(* Logix 5000 project; controller R400_500_XLS vendor 1 type 14 code 216 rev 31.11; software revision 31.01; part 25 of 32 *)
(* tags used below, declared in another part *)
   Abort1 : DINT;   // Not Used
   Alarm : SINT;   // Wait 3 seconds
   AlarmAcked : BOOL;   // Alarm has been acked
   bAlrm : BOOL[64];
   CycExcBuffer : UDT_CYCLE;
   DrainNo : DINT;
   DrnSmp : DINT;
   DRYING : DINT;   // Drying id number
   F1rinse : DINT;   // Not Used
   Fill_Sump : DINT;
   Inj_Time : SINT;   // Time based chemical injection steps
   Last_PwWshRnseTtr : DINT;
   M : DINT[5];   // Memory Bits
   ONS_FC11 : DINT;
   ONS_FC13 : DINT;
   PwExcBuffer : UDT_PW;
   RinseExcBuffer : UDT_RINSE;
   Run : DINT;
   SumpWaterVolume : DINT;   // Sump Water Volume 0 =Low 1= High
   Tmr : TIMER[107];
   Trt_PrWsh : DINT;
   Trt_Rinse : DINT;   // Rinse steps
   Trt_Wsh : DINT;
   WASH_1 : DINT;   // Wash 1 id number
   WASH_5 : DINT;   // Wash 5 id number
   WaterSaved : BOOL;   // Water Saved In Sump (Last Final Rinse Water)
   WshExcBuffer : UDT_WASH;
   bPureWaterFillingAuthorization : BOOL;   // Pure Water Filling Authorization Signal
   DrainExtensionTime : DINT;
   I_Shlf_Sw : BOOL;   // Shelf switch
   I_Smp_Lvl_Hgh : BOOL;   // Sump high level switch
   I_Smp_Lvl_Lw : BOOL;   // Sump low level switch
   msg : BOOL[512];
   PreHeatTime : DINT;
   SumpAlarmFillTime : DINT;
   SumpTemp : REAL;   // Sump temperature in °C
   SumpTempToCool : REAL;   // Sump temperature in °C
   tDelayBeforeFillingAuthAlarm : TIMER;
   tPWClosingDelay : TIMER;
   TreatmentPtr : DINT;
   Unit : Hrdwre;   // Unit Configuration
(* MainProgram, continued *)

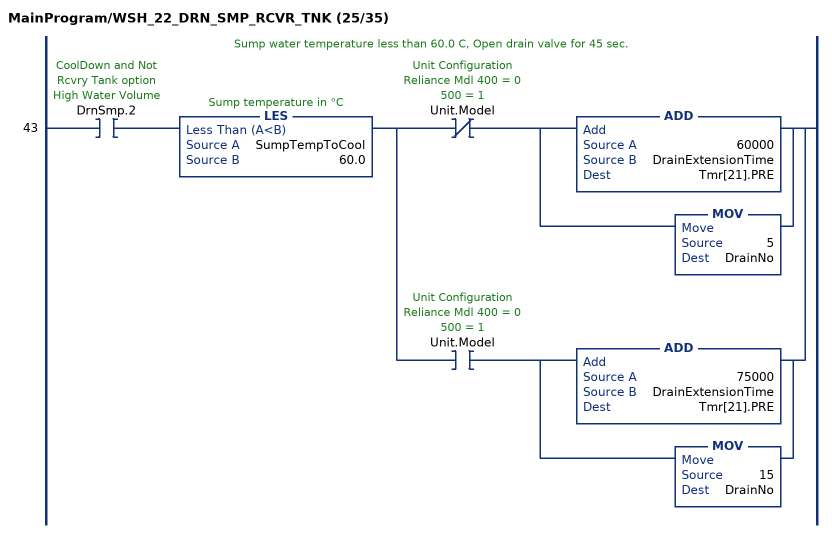
   [picture p501: MainProgram/WSH_22_DRN_SMP_RCVR_TNK rungs 43-43]
   // Sump water temperature less than 60.0 C, Open drain valve for 45 sec.
   43: XIC(DrnSmp.2)LES(SumpTempToCool,60.0)[XIO(Unit.Model) [ADD(60000,DrainExtensionTime,Tmr[21].PRE) ,MOV(5,DrainNo) ] ,XIC(Unit.Model) [ADD(75000,DrainExtensionTime,Tmr[21].PRE) ,MOV(15,DrainNo) ] ];
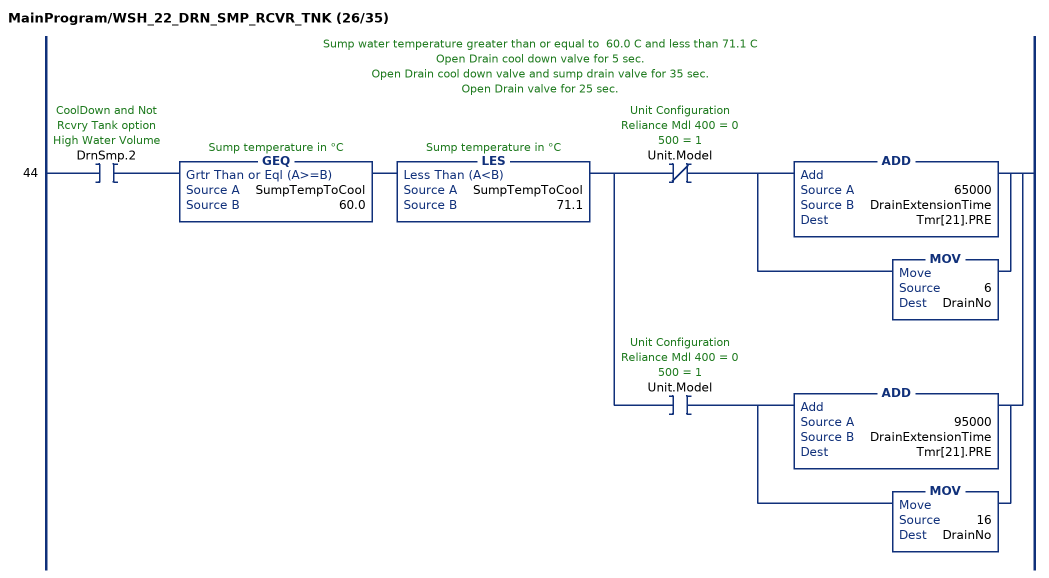
   // Sump water temperature greater than or equal to  60.0 C and less than 71.1 C
   // Open Drain cool down valve for 5 sec.
   // Open Drain cool down valve and sump drain valve for 35 sec.
   // Open Drain valve for 25 sec.
   44: XIC(DrnSmp.2)GEQ(SumpTempToCool,60.0)LES(SumpTempToCool,71.1)[XIO(Unit.Model) [ADD(65000,DrainExtensionTime,Tmr[21].PRE) ,MOV(6,DrainNo) ] ,XIC(Unit.Model) [ADD(95000,DrainExtensionTime,Tmr[21].PRE) ,MOV(16,DrainNo) ] ];
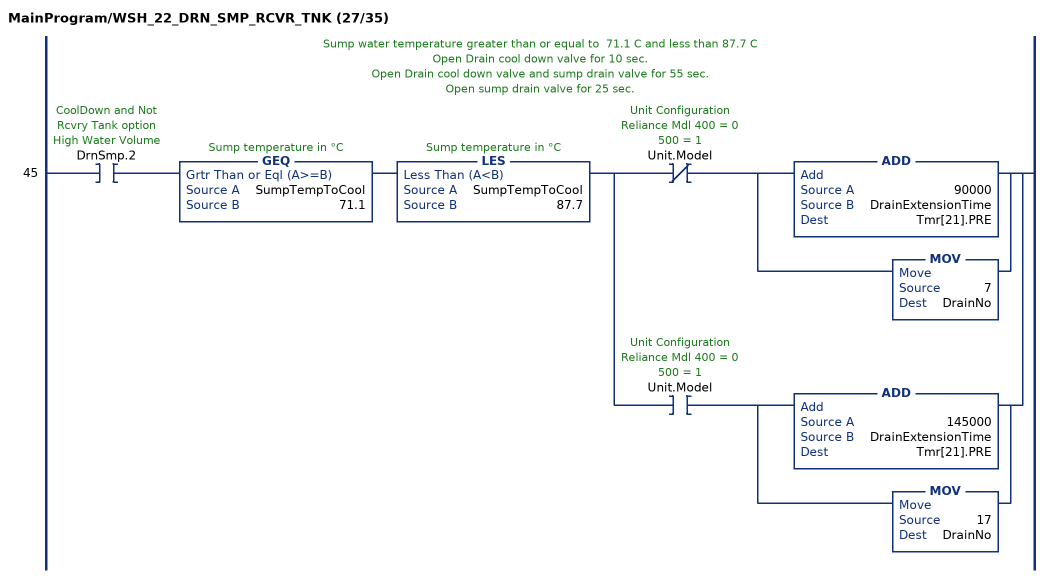
   // Sump water temperature greater than or equal to  71.1 C and less than 87.7 C
   // Open Drain cool down valve for 10 sec.
   // Open Drain cool down valve and sump drain valve for 55 sec.
   // Open sump drain valve for 25 sec.
   45: XIC(DrnSmp.2)GEQ(SumpTempToCool,71.1)LES(SumpTempToCool,87.7)[XIO(Unit.Model) [ADD(90000,DrainExtensionTime,Tmr[21].PRE) ,MOV(7,DrainNo) ] ,XIC(Unit.Model) [ADD(145000,DrainExtensionTime,Tmr[21].PRE) ,MOV(17,DrainNo) ] ];
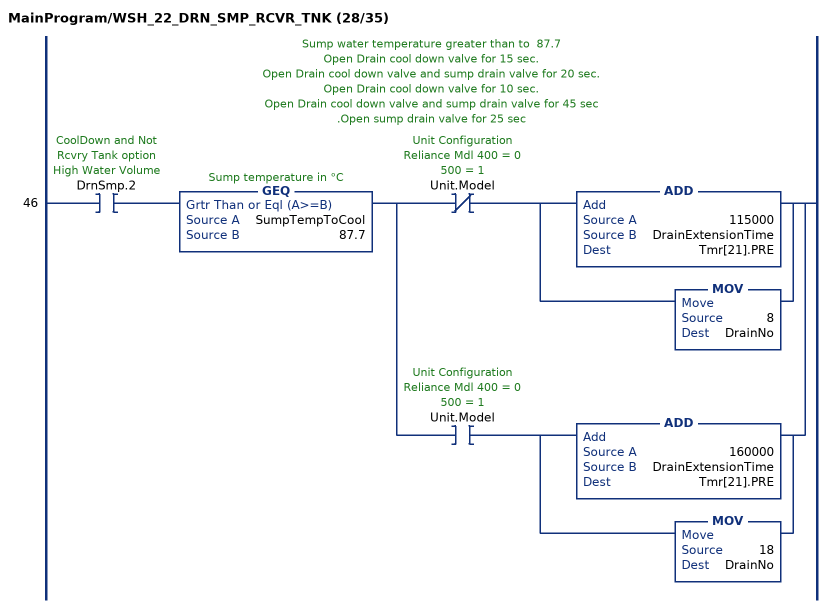
   // Sump water temperature greater than to  87.7
   // Open Drain cool down valve for 15 sec.
   // Open Drain cool down valve and sump drain valve for 20 sec.
   // Open Drain cool down valve for 10 sec.
   // Open Drain cool down valve and sump drain valve for 45 sec
   // .Open sump drain valve for 25 sec
   46: XIC(DrnSmp.2)GEQ(SumpTempToCool,87.7)[XIO(Unit.Model) [ADD(115000,DrainExtensionTime,Tmr[21].PRE) ,MOV(8,DrainNo) ] ,XIC(Unit.Model) [ADD(160000,DrainExtensionTime,Tmr[21].PRE) ,MOV(18,DrainNo) ] ];
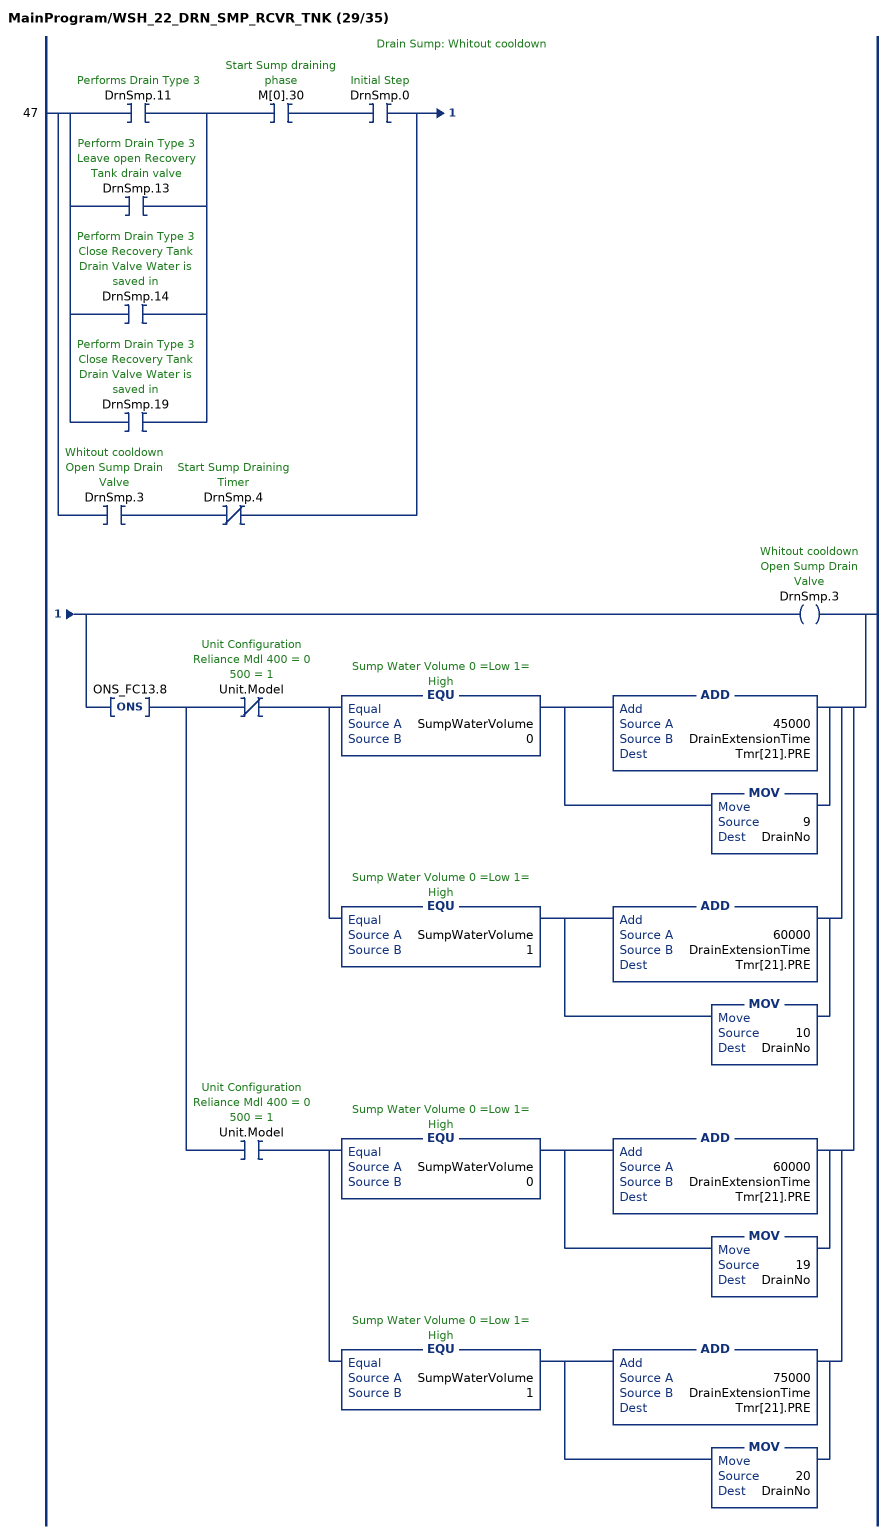
   // Drain Sump: Whitout cooldown
   47: [[XIC(DrnSmp.11) ,XIC(DrnSmp.13) ,XIC(DrnSmp.14) ,XIC(DrnSmp.19) ] XIC(M[0].30) XIC(DrnSmp.0) ,XIC(DrnSmp.3) XIO(DrnSmp.4) ][OTE(DrnSmp.3) ,ONS(ONS_FC13.8) [XIO(Unit.Model) [EQU(SumpWaterVolume,0) [ADD(45000,DrainExtensionTime,Tmr[21].PRE) ,MOV(9,DrainNo) ] ,EQU(SumpWaterVolume,1) [ADD(60000,DrainExtensionTime,Tmr[21].PRE) ,MOV(10,DrainNo) ] ] ,XIC(Unit.Model) [EQU(SumpWaterVolume,0) [ADD(60000,DrainExtensionTime,Tmr[21].PRE) ,MOV(19,DrainNo) ] ,EQU(SumpWaterVolume,1) [ADD(75000,DrainExtensionTime,Tmr[21].PRE) ,MOV(20,DrainNo) ] ] ] ];
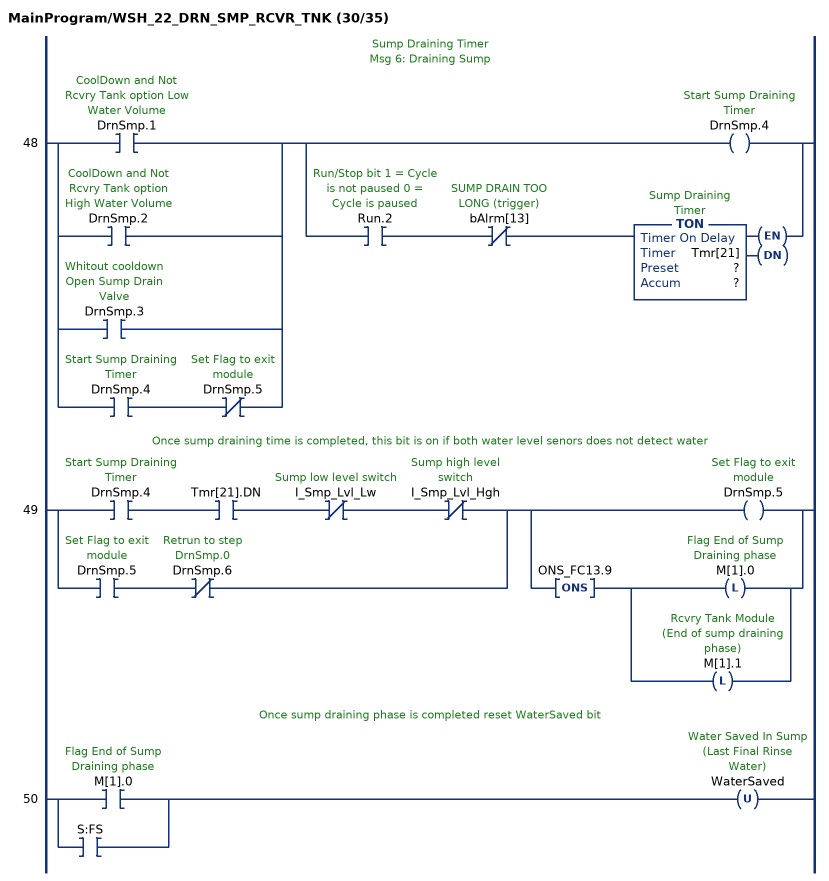
   // Sump Draining Timer
   // Msg 6: Draining Sump
   48: [[XIC(DrnSmp.1) ,XIC(DrnSmp.2) ,XIC(DrnSmp.3) ] ,XIC(DrnSmp.4) XIO(DrnSmp.5) ][OTE(DrnSmp.4) ,XIC(Run.2) XIO(bAlrm[13]) TON(Tmr[21],?,?) ];
   // Once sump draining time is completed, this bit is on if both water level senors does not detect water
   49: [XIC(DrnSmp.4) XIC(Tmr[21].DN) XIO(I_Smp_Lvl_Lw) XIO(I_Smp_Lvl_Hgh) ,XIC(DrnSmp.5) XIO(DrnSmp.6) ][OTE(DrnSmp.5) ,ONS(ONS_FC13.9) [OTL(M[1].0) ,OTL(M[1].1) ] ];
   // Once sump draining phase is completed reset WaterSaved bit
   50: [XIC(M[1].0) ,XIC(S:FS) ]OTU(WaterSaved);
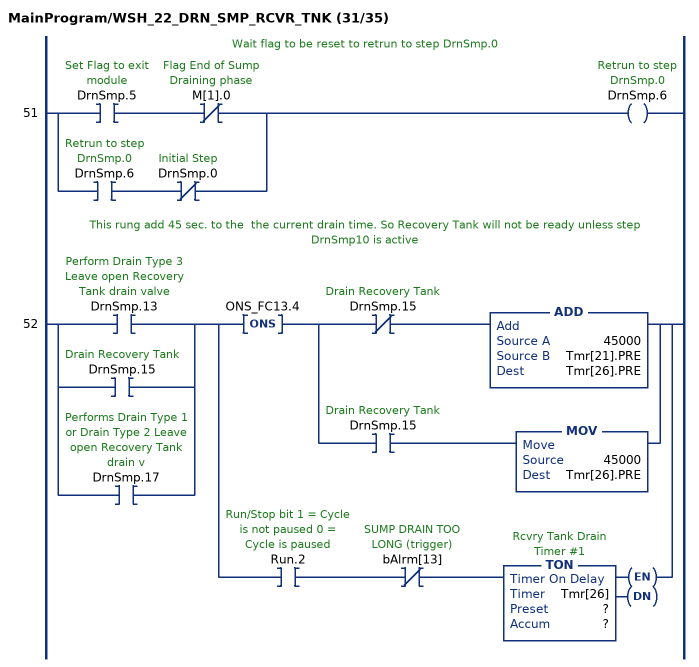
   // Wait flag to be reset to retrun to step DrnSmp.0
   51: [XIC(DrnSmp.5) XIO(M[1].0) ,XIC(DrnSmp.6) XIO(DrnSmp.0) ]OTE(DrnSmp.6);
   // This rung add 45 sec. to the  the current drain time. So Recovery Tank will not be ready unless step DrnSmp10 is active
   52: [XIC(DrnSmp.13) ,XIC(DrnSmp.15) ,XIC(DrnSmp.17) ][ONS(ONS_FC13.4) [XIO(DrnSmp.15) ADD(45000,Tmr[21].PRE,Tmr[26].PRE) ,XIC(DrnSmp.15) MOV(45000,Tmr[26].PRE) ] ,XIC(Run.2) XIO(bAlrm[13]) TON(Tmr[26],?,?) ];
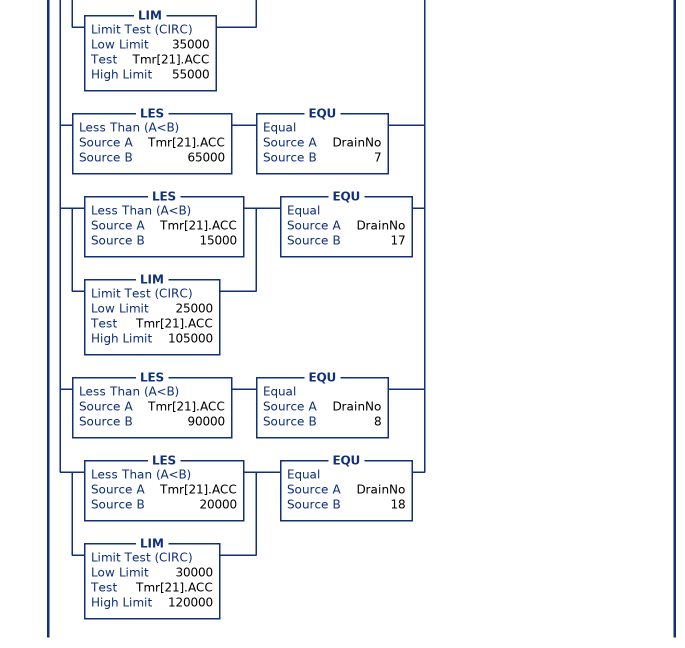
   // Open drain cooldown valve
   53: [LES(Tmr[21].ACC,25000) EQU(DrainNo,2) ,LES(Tmr[21].ACC,35000) EQU(DrainNo,12) ,LES(Tmr[21].ACC,45000) EQU(DrainNo,3) ,[LES(Tmr[21].ACC,15000) ,LIM(25000,Tmr[21].ACC,80000) ] EQU(DrainNo,13) ,LES(Tmr[21].ACC,55000) EQU(DrainNo,4) ,[LES(Tmr[21].ACC,20000) ,LIM(30000,Tmr[21].ACC,90000) ] EQU(DrainNo,14) ,LES(Tmr[21].ACC,40000) EQU(DrainNo,6) ,[LES(Tmr[21].ACC,15000) ,LIM(20000,Tmr[21].ACC,30000) ,LIM(35000,Tmr[21].ACC,55000) ] EQU(DrainNo,16) ,LES(Tmr[21].ACC,65000) EQU(DrainNo,7) ,[LES(Tmr[21].ACC,15000) ,LIM(25000,Tmr[21].ACC,105000) ] EQU(DrainNo,17) ,LES(Tmr[21].ACC,90000) EQU(DrainNo,8) ,[LES(Tmr[21].ACC,20000) ,LIM(30000,Tmr[21].ACC,120000) ] EQU(DrainNo,18) ]XIC(Tmr[21].TT)OTE(DrnSmp.7);
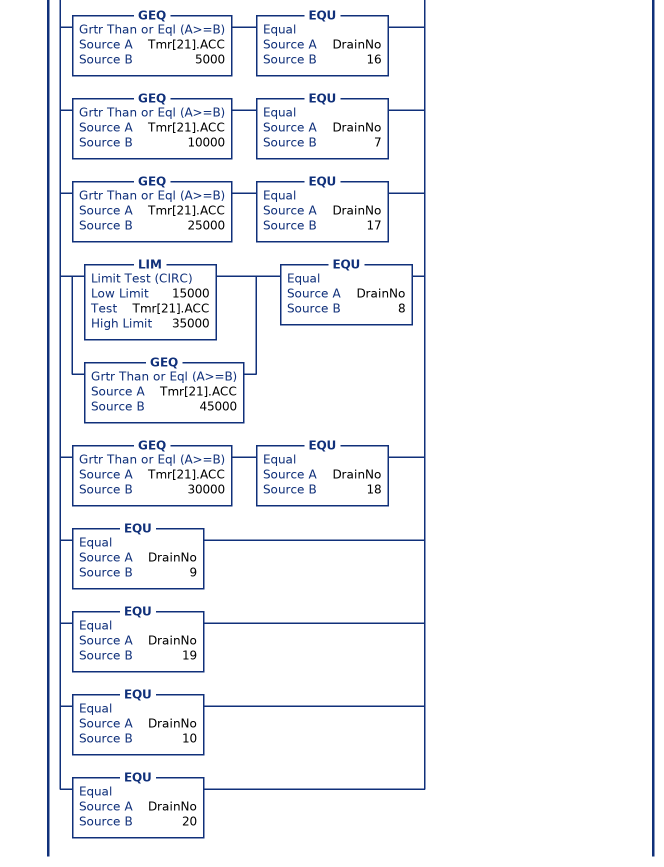
   // Open sump drain valve
   54: [EQU(DrainNo,1) ,EQU(DrainNo,11) ,GEQ(Tmr[21].ACC,5000) EQU(DrainNo,2) ,[LIM(5000,Tmr[21].ACC,15000) ,GEQ(Tmr[21].ACC,20000) ] EQU(DrainNo,12) ,GEQ(Tmr[21].ACC,10000) EQU(DrainNo,3) ,GEQ(Tmr[21].ACC,25000) EQU(DrainNo,13) ,GEQ(Tmr[21].ACC,15000) EQU(DrainNo,4) ,GEQ(Tmr[21].ACC,30000) EQU(DrainNo,14) ,EQU(DrainNo,5) ,EQU(DrainNo,15) ,GEQ(Tmr[21].ACC,5000) EQU(DrainNo,6) ,GEQ(Tmr[21].ACC,5000) EQU(DrainNo,16) ,GEQ(Tmr[21].ACC,10000) EQU(DrainNo,7) ,GEQ(Tmr[21].ACC,25000) EQU(DrainNo,17) ,[LIM(15000,Tmr[21].ACC,35000) ,GEQ(Tmr[21].ACC,45000) ] EQU(DrainNo,8) ,GEQ(Tmr[21].ACC,30000) EQU(DrainNo,18) ,EQU(DrainNo,9) ,EQU(DrainNo,19) ,EQU(DrainNo,10) ,EQU(DrainNo,20) ]XIC(Tmr[21].TT)OTE(DrnSmp.8);
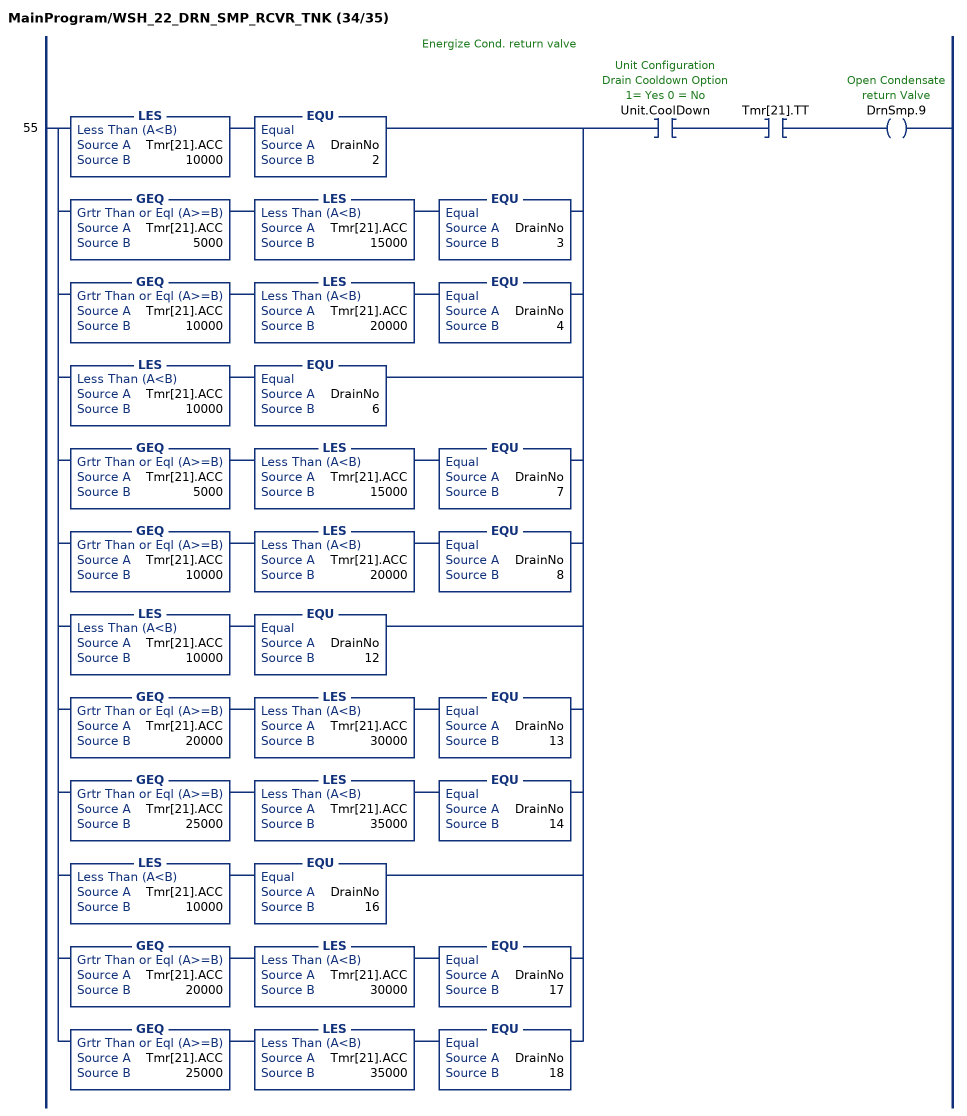
   // Energize Cond. return valve
   55: [LES(Tmr[21].ACC,10000) EQU(DrainNo,2) ,GEQ(Tmr[21].ACC,5000) LES(Tmr[21].ACC,15000) EQU(DrainNo,3) ,GEQ(Tmr[21].ACC,10000) LES(Tmr[21].ACC,20000) EQU(DrainNo,4) ,LES(Tmr[21].ACC,10000) EQU(DrainNo,6) ,GEQ(Tmr[21].ACC,5000) LES(Tmr[21].ACC,15000) EQU(DrainNo,7) ,GEQ(Tmr[21].ACC,10000) LES(Tmr[21].ACC,20000) EQU(DrainNo,8) ,LES(Tmr[21].ACC,10000) EQU(DrainNo,12) ,GEQ(Tmr[21].ACC,20000) LES(Tmr[21].ACC,30000) EQU(DrainNo,13) ,GEQ(Tmr[21].ACC,25000) LES(Tmr[21].ACC,35000) EQU(DrainNo,14) ,LES(Tmr[21].ACC,10000) EQU(DrainNo,16) ,GEQ(Tmr[21].ACC,20000) LES(Tmr[21].ACC,30000) EQU(DrainNo,17) ,GEQ(Tmr[21].ACC,25000) LES(Tmr[21].ACC,35000) EQU(DrainNo,18) ]XIC(Unit.CoolDown)XIC(Tmr[21].TT)OTE(DrnSmp.9);
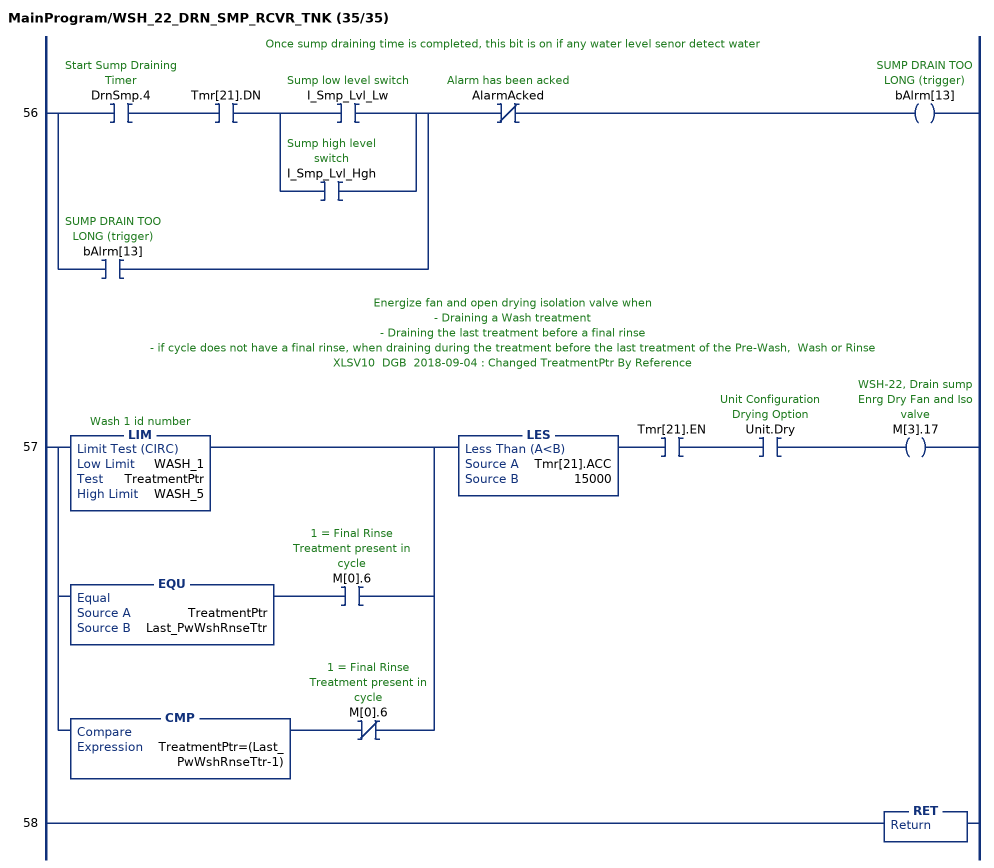
   // Once sump draining time is completed, this bit is on if any water level senor detect water
   56: [XIC(DrnSmp.4) XIC(Tmr[21].DN) [XIC(I_Smp_Lvl_Lw) ,XIC(I_Smp_Lvl_Hgh) ] ,XIC(bAlrm[13]) ]XIO(AlarmAcked)OTE(bAlrm[13]);
   // Energize fan and open drying isolation valve when
   // - Draining a Wash treatment
   // - Draining the last treatment before a final rinse
   // - if cycle does not have a final rinse, when draining during the treatment before the last treatment of the Pre-Wash,  Wash or Rinse
   // XLSV10  DGB  2018-09-04 : Changed TreatmentPtr By Reference
   57: [LIM(WASH_1,TreatmentPtr,WASH_5) ,EQU(TreatmentPtr,Last_PwWshRnseTtr) XIC(M[0].6) ,CMP(TreatmentPtr=(Last_PwWshRnseTtr-1)) XIO(M[0].6) ]LES(Tmr[21].ACC,15000)XIC(Tmr[21].EN)XIC(Unit.Dry)OTE(M[3].17);
   58: RET();
END_ROUTINE

ROUTINE WSH_26_FC11_FILL_SUMP   (* ladder *)
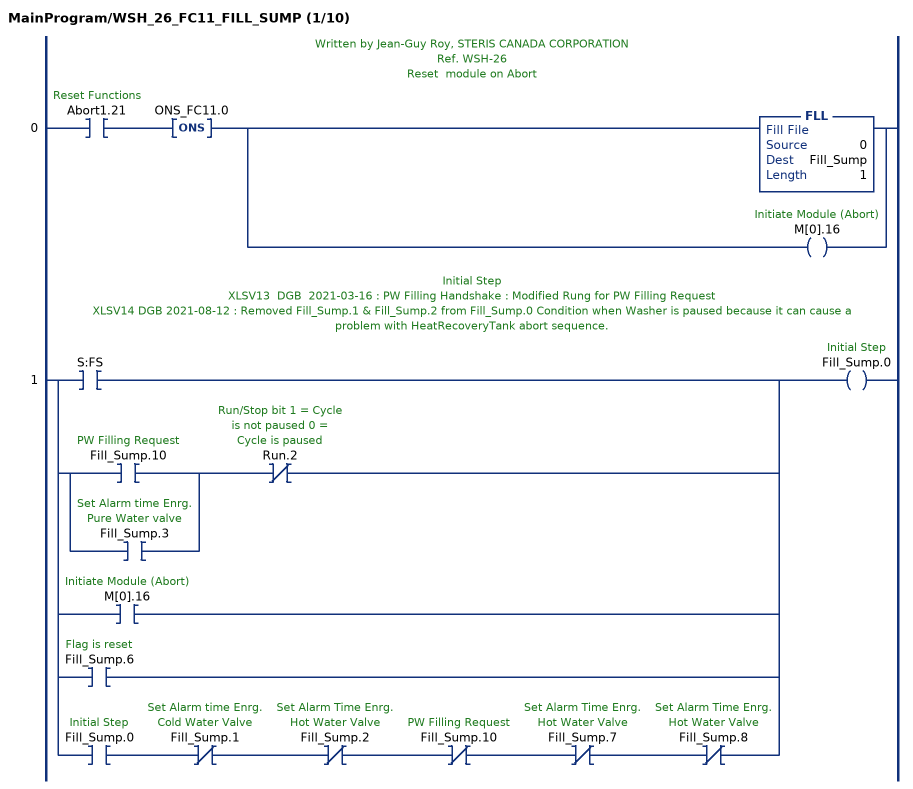
   // Written by Jean-Guy Roy, STERIS CANADA CORPORATION
   // Ref. WSH-26
   // Reset  module on Abort
   0: XIC(Abort1.21)ONS(ONS_FC11.0)[FLL(0,Fill_Sump,1) ,OTE(M[0].16) ];
   // Initial Step
   // XLSV13  DGB  2021-03-16 : PW Filling Handshake : Modified Rung for PW Filling Request
   // XLSV14 DGB 2021-08-12 : Removed Fill_Sump.1 & Fill_Sump.2 from Fill_Sump.0 Condition when Washer is paused because it can cause a problem with HeatRecoveryTank abort sequence.
   1: [XIC(S:FS) ,[XIC(Fill_Sump.10) ,XIC(Fill_Sump.3) ] XIO(Run.2) ,XIC(M[0].16) ,XIC(Fill_Sump.6) ,XIC(Fill_Sump.0) XIO(Fill_Sump.1) XIO(Fill_Sump.2) XIO(Fill_Sump.10) XIO(Fill_Sump.7) XIO(Fill_Sump.8) ]OTE(Fill_Sump.0);
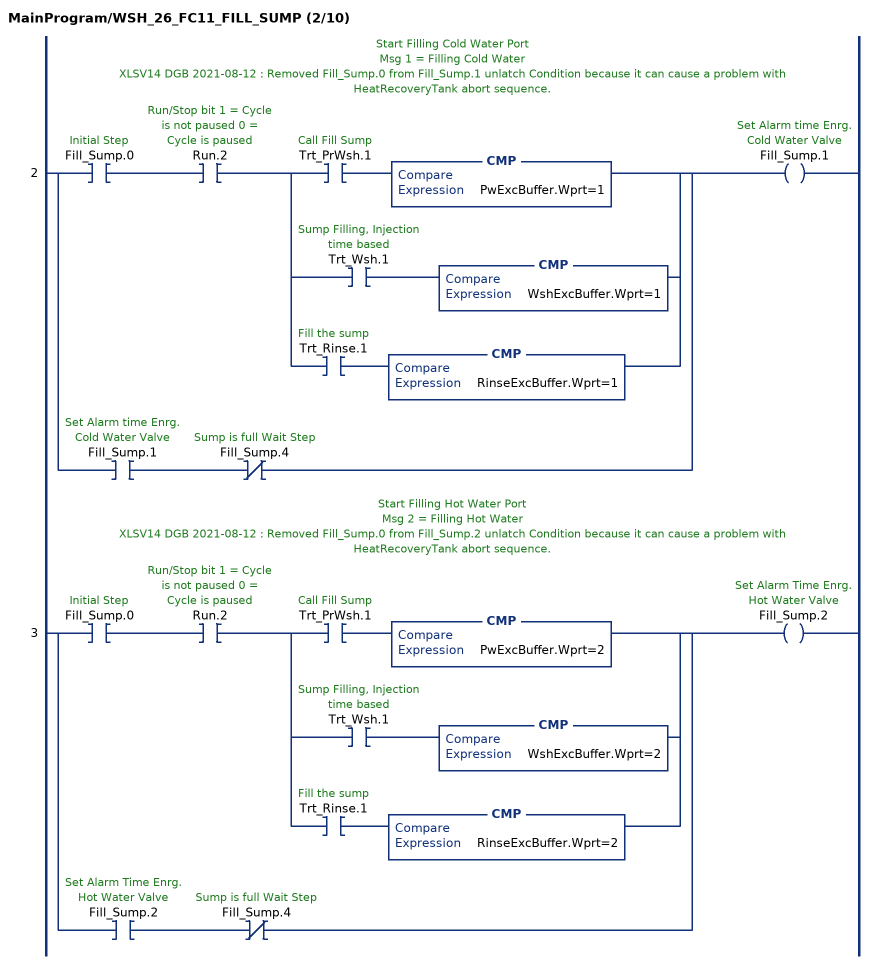
   // Start Filling Cold Water Port
   // Msg 1 = Filling Cold Water
   // XLSV14 DGB 2021-08-12 : Removed Fill_Sump.0 from Fill_Sump.1 unlatch Condition because it can cause a problem with HeatRecoveryTank abort sequence.
   2: [XIC(Fill_Sump.0) XIC(Run.2) [XIC(Trt_PrWsh.1) CMP(PwExcBuffer.Wprt=1) ,XIC(Trt_Wsh.1) CMP(WshExcBuffer.Wprt=1) ,XIC(Trt_Rinse.1) CMP(RinseExcBuffer.Wprt=1) ] ,XIC(Fill_Sump.1) XIO(Fill_Sump.4) ]OTE(Fill_Sump.1);
   // Start Filling Hot Water Port
   // Msg 2 = Filling Hot Water
   // XLSV14 DGB 2021-08-12 : Removed Fill_Sump.0 from Fill_Sump.2 unlatch Condition because it can cause a problem with HeatRecoveryTank abort sequence.
   3: [XIC(Fill_Sump.0) XIC(Run.2) [XIC(Trt_PrWsh.1) CMP(PwExcBuffer.Wprt=2) ,XIC(Trt_Wsh.1) CMP(WshExcBuffer.Wprt=2) ,XIC(Trt_Rinse.1) CMP(RinseExcBuffer.Wprt=2) ] ,XIC(Fill_Sump.2) XIO(Fill_Sump.4) ]OTE(Fill_Sump.2);
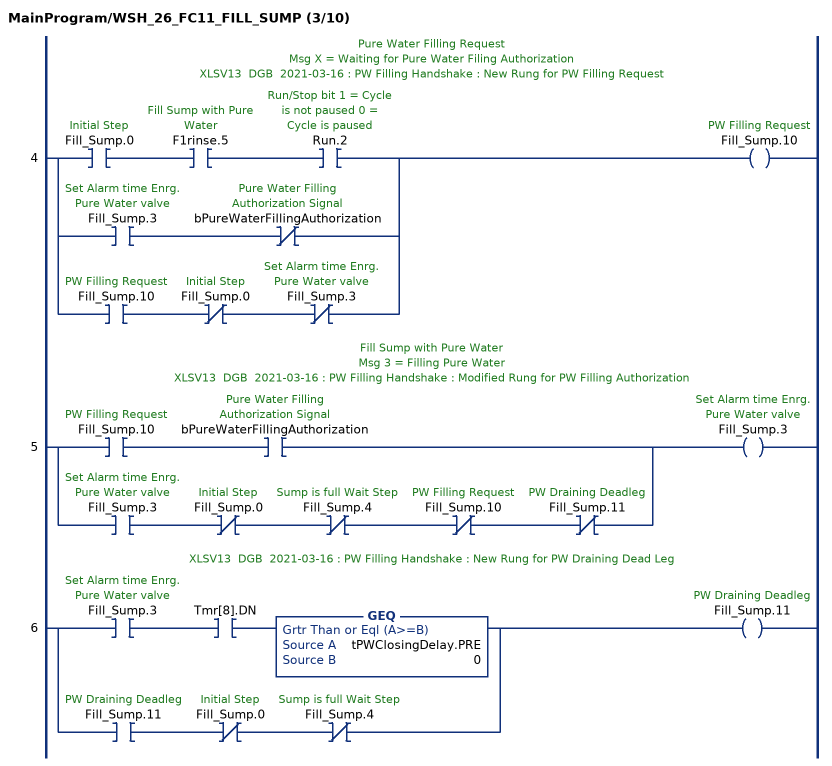
   // Pure Water Filling Request
   // Msg X = Waiting for Pure Water Filing Authorization
   // XLSV13  DGB  2021-03-16 : PW Filling Handshake : New Rung for PW Filling Request
   4: [XIC(Fill_Sump.0) XIC(F1rinse.5) XIC(Run.2) ,XIC(Fill_Sump.3) XIO(bPureWaterFillingAuthorization) ,XIC(Fill_Sump.10) XIO(Fill_Sump.0) XIO(Fill_Sump.3) ]OTE(Fill_Sump.10);
   // Fill Sump with Pure Water
   // Msg 3 = Filling Pure Water
   // XLSV13  DGB  2021-03-16 : PW Filling Handshake : Modified Rung for PW Filling Authorization
   5: [XIC(Fill_Sump.10) XIC(bPureWaterFillingAuthorization) ,XIC(Fill_Sump.3) XIO(Fill_Sump.0) XIO(Fill_Sump.4) XIO(Fill_Sump.10) XIO(Fill_Sump.11) ]OTE(Fill_Sump.3);
   // XLSV13  DGB  2021-03-16 : PW Filling Handshake : New Rung for PW Draining Dead Leg
   6: [XIC(Fill_Sump.3) XIC(Tmr[8].DN) GEQ(tPWClosingDelay.PRE,0) ,XIC(Fill_Sump.11) XIO(Fill_Sump.0) XIO(Fill_Sump.4) ]OTE(Fill_Sump.11);
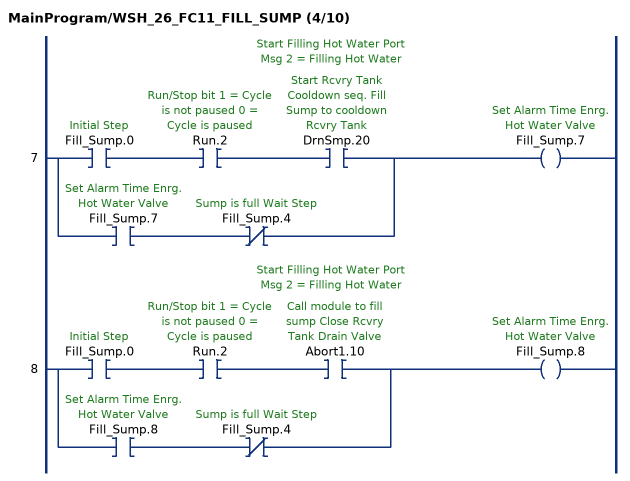
   // Start Filling Hot Water Port
   // Msg 2 = Filling Hot Water
   7: [XIC(Fill_Sump.0) XIC(Run.2) XIC(DrnSmp.20) ,XIC(Fill_Sump.7) XIO(Fill_Sump.4) ]OTE(Fill_Sump.7);
   // Start Filling Hot Water Port
   // Msg 2 = Filling Hot Water
   8: [XIC(Fill_Sump.0) XIC(Run.2) XIC(Abort1.10) ,XIC(Fill_Sump.8) XIO(Fill_Sump.4) ]OTE(Fill_Sump.8);
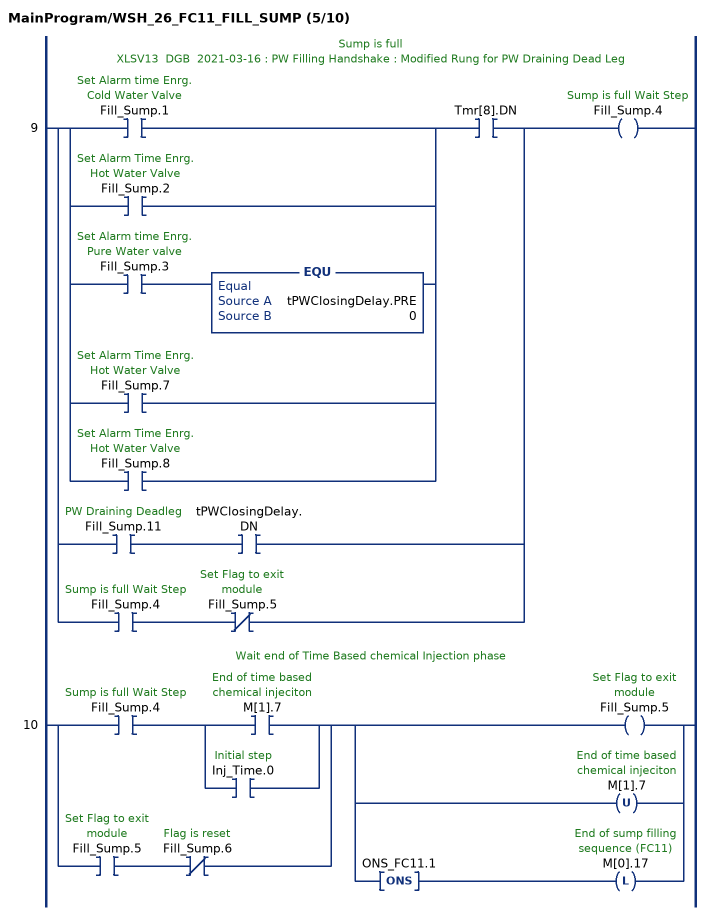
   // Sump is full
   // XLSV13  DGB  2021-03-16 : PW Filling Handshake : Modified Rung for PW Draining Dead Leg
   9: [[XIC(Fill_Sump.1) ,XIC(Fill_Sump.2) ,XIC(Fill_Sump.3) EQU(tPWClosingDelay.PRE,0) ,XIC(Fill_Sump.7) ,XIC(Fill_Sump.8) ] XIC(Tmr[8].DN) ,XIC(Fill_Sump.11) XIC(tPWClosingDelay.DN) ,XIC(Fill_Sump.4) XIO(Fill_Sump.5) ]OTE(Fill_Sump.4);
   // Wait end of Time Based chemical Injection phase
   10: [XIC(Fill_Sump.4) [XIC(M[1].7) ,XIC(Inj_Time.0) ] ,XIC(Fill_Sump.5) XIO(Fill_Sump.6) ][OTE(Fill_Sump.5) ,OTU(M[1].7) ,ONS(ONS_FC11.1) OTL(M[0].17) ];
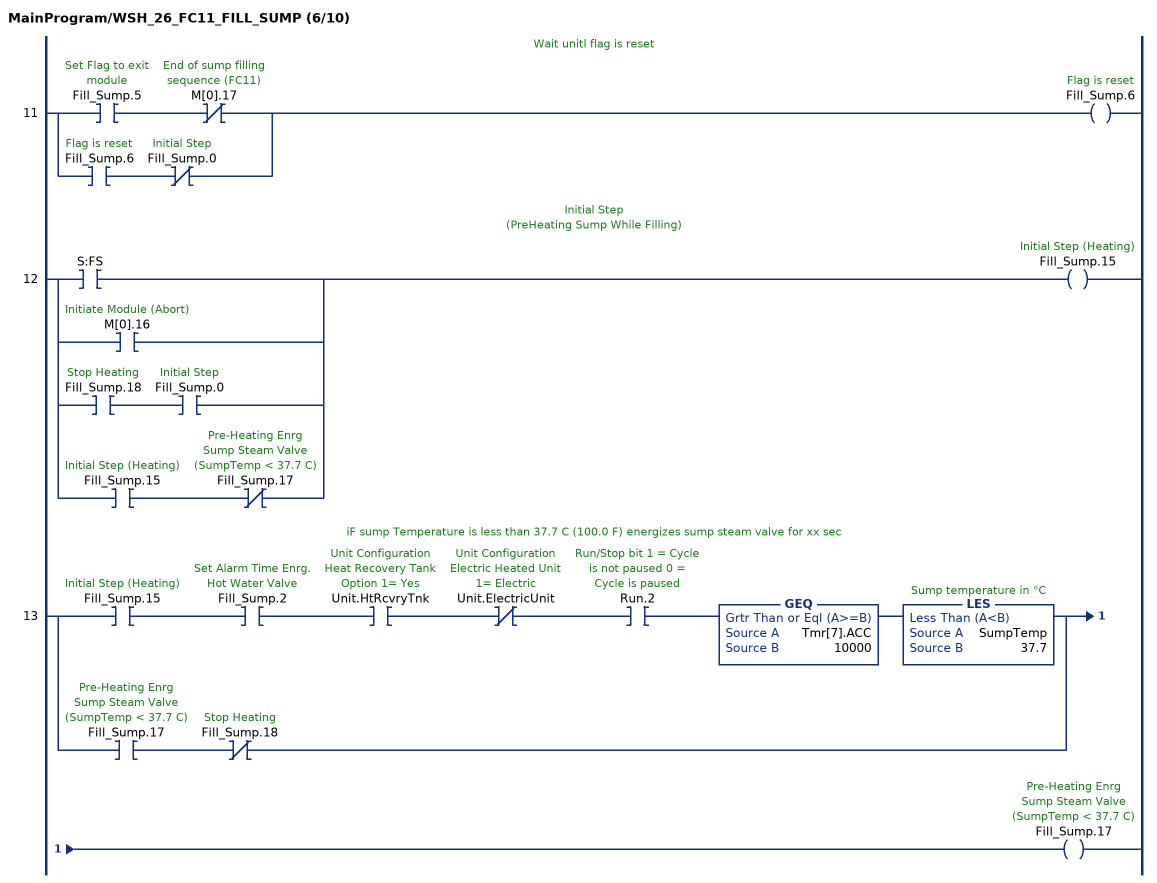
   // Wait unitl flag is reset
   11: [XIC(Fill_Sump.5) XIO(M[0].17) ,XIC(Fill_Sump.6) XIO(Fill_Sump.0) ]OTE(Fill_Sump.6);
   // Initial Step
   // (PreHeating Sump While Filling)
   12: [XIC(S:FS) ,XIC(M[0].16) ,XIC(Fill_Sump.18) XIC(Fill_Sump.0) ,XIC(Fill_Sump.15) XIO(Fill_Sump.17) ]OTE(Fill_Sump.15);
   // iF sump Temperature is less than 37.7 C (100.0 F) energizes sump steam valve for xx sec
   13: [XIC(Fill_Sump.15) XIC(Fill_Sump.2) XIC(Unit.HtRcvryTnk) XIO(Unit.ElectricUnit) XIC(Run.2) GEQ(Tmr[7].ACC,10000) LES(SumpTemp,37.7) ,XIC(Fill_Sump.17) XIO(Fill_Sump.18) ]OTE(Fill_Sump.17);
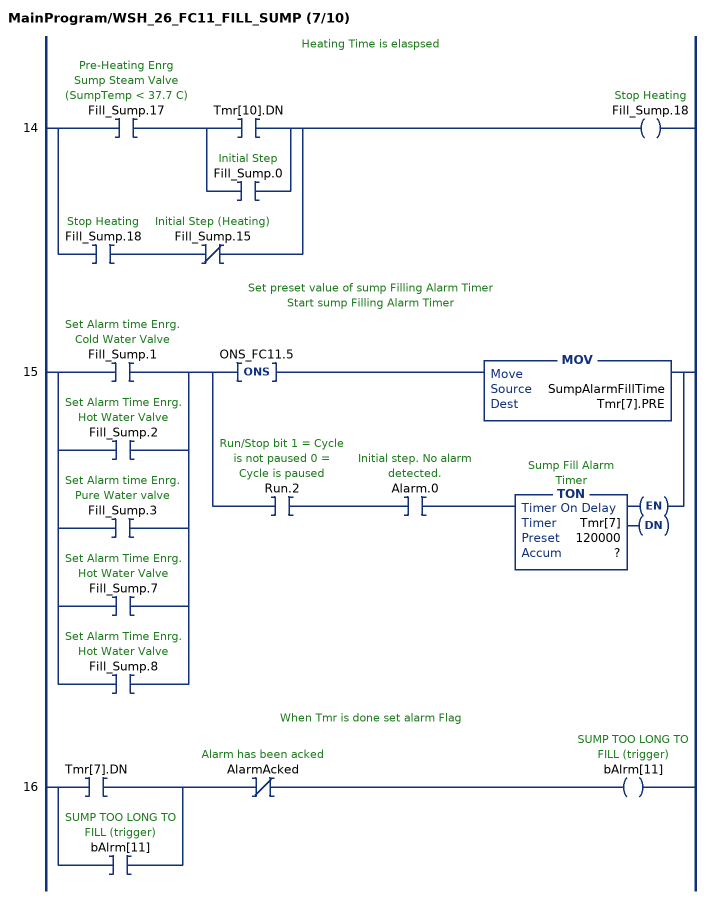
   // Heating Time is elaspsed
   14: [XIC(Fill_Sump.17) [XIC(Tmr[10].DN) ,XIC(Fill_Sump.0) ] ,XIC(Fill_Sump.18) XIO(Fill_Sump.15) ]OTE(Fill_Sump.18);
   // Set preset value of sump Filling Alarm Timer
   // Start sump Filling Alarm Timer
   15: [XIC(Fill_Sump.1) ,XIC(Fill_Sump.2) ,XIC(Fill_Sump.3) ,XIC(Fill_Sump.7) ,XIC(Fill_Sump.8) ][ONS(ONS_FC11.5) MOV(SumpAlarmFillTime,Tmr[7].PRE) ,XIC(Run.2) XIC(Alarm.0) TON(Tmr[7],?,?) ];
   // When Tmr is done set alarm Flag
   16: [XIC(Tmr[7].DN) ,XIC(bAlrm[11]) ]XIO(AlarmAcked)OTE(bAlrm[11]);
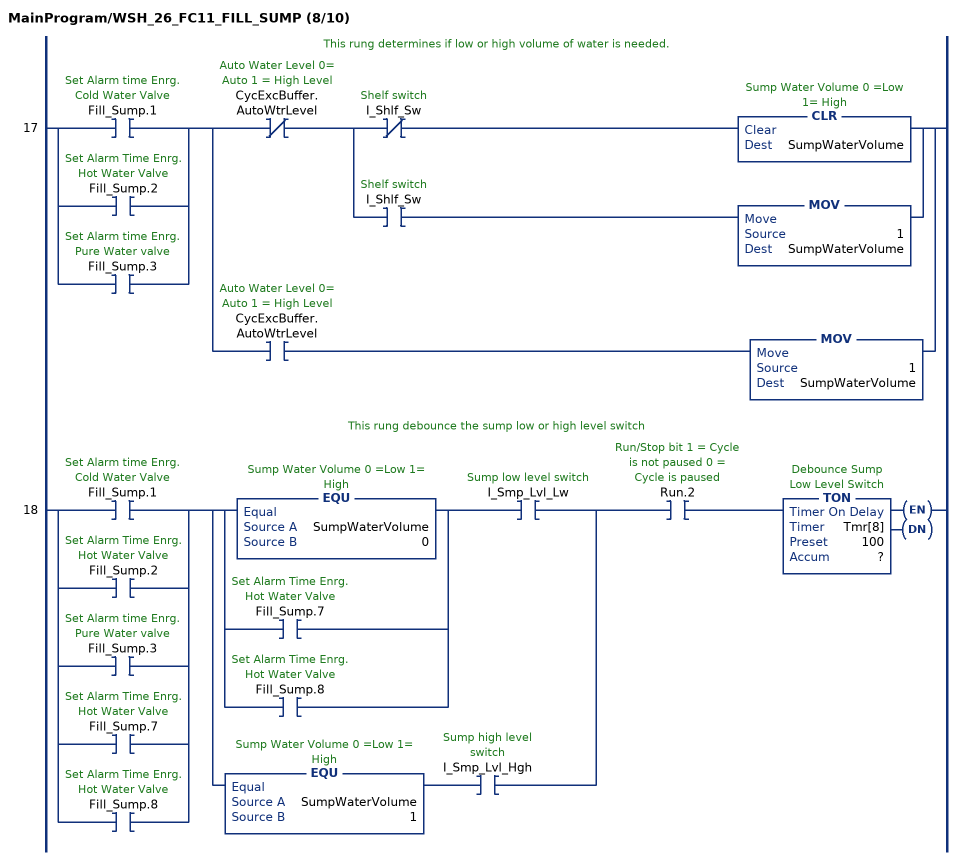
   // This rung determines if low or high volume of water is needed.
   17: [XIC(Fill_Sump.1) ,XIC(Fill_Sump.2) ,XIC(Fill_Sump.3) ][XIO(CycExcBuffer.AutoWtrLevel) [XIO(I_Shlf_Sw) CLR(SumpWaterVolume) ,XIC(I_Shlf_Sw) MOV(1,SumpWaterVolume) ] ,XIC(CycExcBuffer.AutoWtrLevel) MOV(1,SumpWaterVolume) ];
   // This rung debounce the sump low or high level switch
   18: [XIC(Fill_Sump.1) ,XIC(Fill_Sump.2) ,XIC(Fill_Sump.3) ,XIC(Fill_Sump.7) ,XIC(Fill_Sump.8) ][[EQU(SumpWaterVolume,0) ,XIC(Fill_Sump.7) ,XIC(Fill_Sump.8) ] XIC(I_Smp_Lvl_Lw) ,EQU(SumpWaterVolume,1) XIC(I_Smp_Lvl_Hgh) ]XIC(Run.2)TON(Tmr[8],?,?);
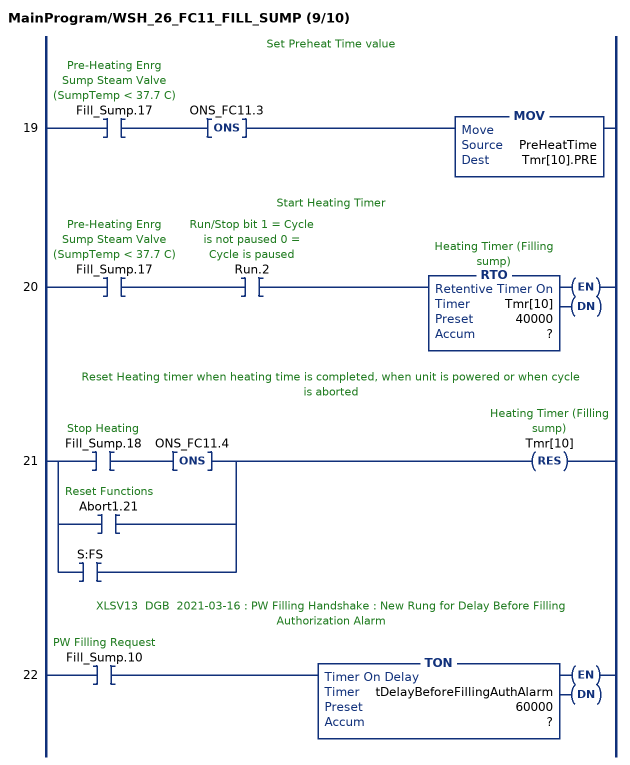
   // Set Preheat Time value
   19: XIC(Fill_Sump.17)ONS(ONS_FC11.3)MOV(PreHeatTime,Tmr[10].PRE);
   // Start Heating Timer
   20: XIC(Fill_Sump.17)XIC(Run.2)RTO(Tmr[10],?,?);
   // Reset Heating timer when heating time is completed, when unit is powered or when cycle is aborted
   21: [XIC(Fill_Sump.18) ONS(ONS_FC11.4) ,XIC(Abort1.21) ,XIC(S:FS) ]RES(Tmr[10]);
   // XLSV13  DGB  2021-03-16 : PW Filling Handshake : New Rung for Delay Before Filling Authorization Alarm
   22: XIC(Fill_Sump.10)TON(tDelayBeforeFillingAuthAlarm,?,?);
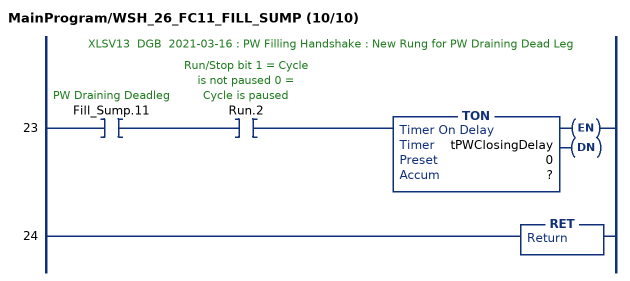
   // XLSV13  DGB  2021-03-16 : PW Filling Handshake : New Rung for PW Draining Dead Leg
   23: XIC(Fill_Sump.11)XIC(Run.2)TON(tPWClosingDelay,?,?);
   24: RET();
END_ROUTINE
